(* IEC 61131-3 sources: llm-plc-st-eval/data/calibracion/qwen2.5-coder_14b/B1/few_shot, 3 files *)

(* ---- ejec_1.st ---- *)
FUNCTION_BLOCK FB_Motor
VAR_INPUT
    btnMarcha : BOOL; (* Boton de marcha *)
    btnParo : BOOL; (* Boton de paro *)
    btnEmerg : BOOL; (* Boton de emergencia *)
END_VAR
VAR_OUTPUT
    motorOn : BOOL; (* Estado del motor *)
END_VAR
VAR
    motorStart : BOOL; (* Bandera de arranque *)
    motorStop : BOOL; (* Bandera de paro *)
    emergStop : BOOL; (* Bandera de paro de emergencia *)
END_VAR

(* Control de arranque y paro del motor *)
motorStart := btnMarcha AND NOT motorStop AND NOT emergStop;
motorStop := btnParo OR emergStop;
emergStop := btnEmerg;

(* Actualizar el estado del motor *)
IF motorStart THEN
    motorOn := TRUE;
ELSIF motorStop THEN
    motorOn := FALSE;
END_IF;
END_FUNCTION_BLOCK

(* ---- ejec_2.st ---- *)
FUNCTION_BLOCK FB_Motor
VAR_INPUT
    btnMarcha : BOOL; (* Boton de marcha *)
    btnParo : BOOL; (* Boton de paro *)
    btnEmerg : BOOL; (* Boton de emergencia *)
END_VAR
VAR_OUTPUT
    motorOn : BOOL; (* Estado del motor *)
END_VAR
VAR
    estadoEmergencia : BOOL; (* Estado de emergencia *)
END_VAR

(* Control de arranque y paro del motor *)
IF btnEmerg THEN
    estadoEmergencia := TRUE;
    motorOn := FALSE;
ELSIF estadoEmergencia THEN
    motorOn := FALSE;
ELSIF btnParo THEN
    motorOn := FALSE;
ELSIF btnMarcha THEN
    motorOn := TRUE;
END_IF;
END_FUNCTION_BLOCK

(* ---- ejec_3.st ---- *)
FUNCTION_BLOCK FB_Motor
VAR_INPUT
    btnMarcha : BOOL; (* Boton de marcha *)
    btnParo : BOOL; (* Boton de paro *)
    btnEmerg : BOOL; (* Boton de emergencia *)
END_VAR
VAR_OUTPUT
    motorOn : BOOL; (* Motor encendido *)
END_VAR
VAR
    motorStarted : BOOL; (* Bandera para indicar si el motor ha sido arrancado *)
END_VAR

(* Arranque del motor *)
IF btnMarcha AND NOT motorStarted THEN
    motorStarted := TRUE;
    motorOn := TRUE;
END_IF;

(* Paro del motor *)
IF btnParo OR btnEmerg THEN
    motorStarted := FALSE;
    motorOn := FALSE;
END_IF;

(* Mantener el motor encendido después de arrancarlo *)
IF motorStarted THEN
    motorOn := TRUE;
END_IF;

END_FUNCTION_BLOCK
